TYPE "ST_ConfigPage"
VERSION : 0.1
   STRUCT
      Revision : UDInt;
      PageIndex : Int;
      PageCount : Int;
      EntryCount : Int;
      Entries : Array[1..16] of "ST_ConfigEntry";
   END_STRUCT;

END_TYPE

